# EPICS substitutions: iocs/rr/iocBoot/iocrr/motorSim.substitutions
file "$(MOTOR)/db/asyn_motor_model2.db"
{
pattern
{N,        M,  ADDR,        DESC,  EGU,  DIR,  VELO,  VBAS,  ACCL,  BDST,  BVEL,  BACC,  MRES,  PREC,  DHLM,  DLLM,  INIT}
{1,  "m$(N)",     0,  "$(P)$(M)",   deg,  Pos,   30,     0,    .2,     0,     1,    .2,  0.01,     5,   1e6,  -1e6,    ""}
{2,  "m$(N)",     1,  "$(P)$(M)",   deg,  Pos,   30,     0,    .2,     0,     1,    .2,  0.01,     5,   1e6,  -1e6,    ""}
}
